Fanuc KAREL source: NC0091.KL

-- PROVISIONAL review KL for V940-1; original PC SHA256 57149644955d8b491b5bef8728e3006a14cdb852eaf33b75f58206545ba73da8
-- Incomplete behavior may be omitted. Consult companion uncertainty JSON. Do not deploy.
PROGRAM NC0091
%NOLOCKGROUP
-- UNRESOLVED_LOCAL_POOL 6 cells at code offset 3; source declarations unknown
-- DIRECT_LOCAL_WORD_ACCESS alone does not prove INTEGER, REAL, or BOOLEAN
BEGIN
  -- V9_OWNER_INTERVAL_HINT [23,247),[45,216),[67,185),[89,154),[111,123); structural only; source/VM held
  -- V9_FOOTER_20_HINT 5 numerical footer links; VM transfer unproved
  -- UNRESOLVED_PC offsets 0-8; opcodes 2B,2C,7B
  -- UNRESOLVED_PC offsets 13-20; opcodes 9D,23
  -- UNRESOLVED_PC offsets 25-38; opcodes 21,9D,57,79
  -- UNRESOLVED_PC offsets 43-60; opcodes 21,40,41,42
  -- UNRESOLVED_PC offsets 65-94; opcodes 9D,23,9E,2E,22,7A
  -- UNRESOLVED_PC offsets 99-116; opcodes 21,2E,59,79
  -- UNRESOLVED_PC offsets 121-134; opcodes 21,9D,57,79
  -- UNRESOLVED_PC offsets 139-156; opcodes 21,40,41,42
  -- UNRESOLVED_PC offsets 161-190; opcodes 9D,23,9E,2E,22,7A
  -- UNRESOLVED_PC offsets 195-212; opcodes 21,2E,59,79
  -- UNRESOLVED_PC offsets 217-230; opcodes 21,9D,57,79
  -- UNRESOLVED_PC offsets 235-252; opcodes 21,40,41,42
  -- UNRESOLVED_PC offsets 257-286; opcodes 9D,23,9E,2E,22,7A
  -- UNRESOLVED_PC offsets 291-308; opcodes 21,2E,59,79
  -- UNRESOLVED_PC offsets 313-326; opcodes 21,9D,57,79
  -- UNRESOLVED_PC offsets 331-348; opcodes 21,40,41,42
  -- UNRESOLVED_PC offsets 353-382; opcodes 9D,23,9E,2E,22,7A
  -- UNRESOLVED_PC offsets 387-404; opcodes 21,2E,59,79
  -- UNRESOLVED_PC offsets 409-422; opcodes 21,9D,57,79
  -- UNRESOLVED_PC offsets 427-444; opcodes 21,40,41,42
  -- UNRESOLVED_PC offsets 449-478; opcodes 9D,23,9E,2E,22,7A
  -- UNRESOLVED_PC offsets 483-500; opcodes 21,2E,59,79
  -- UNRESOLVED_PC offsets 505-519; opcodes 21,9D,52,23
  -- UNRESOLVED_PC offsets 524-529; opcodes 7A
  -- UNRESOLVED_PC offsets 534-565; opcodes 20,2C,23,7A,40,41,42
  -- UNRESOLVED_PC offsets 570-594; opcodes 21,2E,52,23,7A,43
  -- UNRESOLVED_PC offsets 599-617; opcodes 21,2E,52,23
  -- UNRESOLVED_PC offsets 627-632; opcodes 7A
  -- UNRESOLVED_PC offsets 637-655; opcodes 21,2E,52,23
  -- UNRESOLVED_PC offsets 665-670; opcodes 7A
  -- UNRESOLVED_PC offsets 675-706; opcodes 20,2C,23,7A,40,41,42
  -- UNRESOLVED_PC offsets 711-735; opcodes 21,2E,52,23,7A,43
  -- UNRESOLVED_PC offsets 740-758; opcodes 21,2E,52,23
  -- UNRESOLVED_PC offsets 768-773; opcodes 7A
  -- UNRESOLVED_PC offsets 778-796; opcodes 21,2E,52,23
  -- UNRESOLVED_PC offsets 806-811; opcodes 7A
  -- UNRESOLVED_PC offsets 816-847; opcodes 20,2C,23,7A,40,41,42
  -- UNRESOLVED_PC offsets 852-876; opcodes 21,2E,52,23,7A,43
  -- UNRESOLVED_PC offsets 881-899; opcodes 21,2E,52,23
  -- UNRESOLVED_PC offsets 909-914; opcodes 7A
  -- UNRESOLVED_PC offsets 919-937; opcodes 21,2E,52,23
  -- UNRESOLVED_PC offsets 947-952; opcodes 7A
  -- UNRESOLVED_PC offsets 957-988; opcodes 20,2C,23,7A,40,41,42
  -- UNRESOLVED_PC offsets 993-1017; opcodes 21,2E,52,23,7A,43
  -- UNRESOLVED_PC offsets 1022-1040; opcodes 21,2E,52,23
  -- UNRESOLVED_PC offsets 1050-1055; opcodes 7A
  -- UNRESOLVED_PC offsets 1060-1078; opcodes 21,2E,52,23
  -- UNRESOLVED_PC offsets 1088-1093; opcodes 7A
  -- UNRESOLVED_PC offsets 1098-1129; opcodes 20,2C,23,7A,40,41,42
  -- UNRESOLVED_PC offsets 1134-1158; opcodes 21,2E,52,23,7A,43
  -- UNRESOLVED_PC offsets 1163-1181; opcodes 21,2E,52,23
  -- UNRESOLVED_PC offsets 1191-1196; opcodes 7A
  -- UNRESOLVED_PC offsets 1201-1219; opcodes 21,2E,52,23
  -- UNRESOLVED_PC offsets 1229-1233; opcodes 7F
  -- UNRESOLVED_PC offsets 1238-1242; opcodes 27,AA
  -- UNRESOLVED_PC offsets 1247-1251; opcodes 7F
END NC0091
